# EPICS autosave request: iocs/ad/pva-driver-ioc/auto_settings.req
file "pvaDriver_settings.req",      P=$(P),  R=cam1:
file "NDStdArrays_settings.req",    P=$(P),  R=image1:
file "commonPlugin_settings.req",   P=$(P)
